SUBAPPLICATION StringValue_TO_NVS (* String-VT-Wert einlesen und in NVS speichern (generisch). *)
  (* Standard: 61499-2 *)
  (* Version 1.0, 2026-09-09, Franz Höpfinger, Meisterschulen am Ostbahnhof, Ausgelagert aus Uebung_012m_sub zur Wiederverwendung. *)
  PACKAGE MyLib::sys;
  IMPORT isobus::UT::Q::const::IDs::ID_NULL;
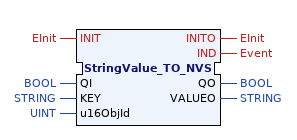
  EVENT_INPUT
    INIT : EInit; (* Initialization Request *)
  END_EVENT
  EVENT_OUTPUT
    INITO : EInit; (* Initialization Confirm *)
    IND;
  END_EVENT
  VAR_INPUT
    QI : BOOL := TRUE; (* Quality Input - TRUE to enable service *)
    KEY : STRING; (* Key name. *)
    u16ObjId : UINT := ID_NULL;
  END_VAR
  VAR_OUTPUT
    QO : BOOL; (* Quality Output - TRUE if service executed successfully *)
    VALUEO : STRING;
  END_VAR
  FBS
    StringValue_IS : isobus::UT::io::StringValue::StringValue_IS;
    NVS : logiBUS::storage::esp32_nvs::NVS(DEFAULT_VALUE := STRING#'');
    Q_StringValue : isobus::UT::Q::Q_StringValue;
    AND_QO : iec61131::booleanOperators::AND_BOOL_3;
  END_FBS
  EVENT_CONNECTIONS
    StringValue_IS.IND TO NVS.SET;
    NVS.SETO TO IND;
    NVS.GETO TO Q_StringValue.REQ;
    NVS.GETO TO IND;
    NVS.INITO TO NVS.GET;
    INIT TO Q_StringValue.INIT;
    Q_StringValue.INITO TO StringValue_IS.INIT;
    StringValue_IS.INITO TO NVS.INIT;
    NVS.INITO TO INITO;
    NVS.INITO TO AND_QO.REQ;
  END_CONNECTIONS
  DATA_CONNECTIONS
    StringValue_IS.IN TO NVS.VALUE;
    u16ObjId TO Q_StringValue.u16ObjId;
    KEY TO NVS.KEY;
    NVS.VALUEO TO Q_StringValue.pau8String;
    NVS.VALUEO TO VALUEO;
    u16ObjId TO StringValue_IS.u16ObjId;
    QI TO Q_StringValue.QI;
    QI TO StringValue_IS.QI;
    QI TO NVS.QI;
    Q_StringValue.QO TO AND_QO.IN1;
    StringValue_IS.QO TO AND_QO.IN2;
    NVS.QO TO AND_QO.IN3;
    AND_QO.OUT TO QO;
  END_CONNECTIONS
END_SUBAPPLICATION
